{region 'Documentation'}
(*!
<summary>Check that IN is inside the inclusive StartTime..EndTime interval.</summary>
<description>

StartTime &gt; EndTime reports Error during active evaluation; equal bounds are
valid.

</description>
*)
{endregion}
FUNCTION_BLOCK AssertInTimespan_DT EXTENDS AssertionBase
VAR_INPUT
    IN : DT; //! Actual value checked or observed by this Assertion.
    StartTime : DT; //! Inclusive start of the time span; must not exceed EndTime.
    EndTime : DT; //! Inclusive end of the time span; must not precede StartTime.
END_VAR

SUPER^();

{region 'Documentation'}
(*!
<summary>Evaluate the typed temporal relation and report higher-priority errors first.</summary>
*)
{endregion}
METHOD PROTECTED Assert
VAR
    Message : STRING(GVL_Constants.MessageLength);
    StartTimeText : STRING(GVL_Constants.AssertionValueLength);
    EndTimeText : STRING(GVL_Constants.AssertionValueLength);
    ActualText : STRING(GVL_Constants.AssertionValueLength);
END_VAR
IF NOT EvaluationActive THEN
    RETURN;
END_IF;

IF Result = E_Result.Error THEN
    RETURN;
END_IF;

IF StartTime > EndTime THEN
    StartTimeText := DT_TO_STRING(StartTime);
    EndTimeText := DT_TO_STRING(EndTime);
    Message := CONCAT('Assertion error: start time exceeds end time. StartTime = ',
        StartTimeText);
    Message := CONCAT(Message, ', EndTime = ');
    Message := CONCAT(Message, EndTimeText);
    Message := CONCAT(Message, '.');
    Error(Message := Message);
    RETURN;
END_IF;

IF Result = E_Result.Failed THEN
    RETURN;
END_IF;

IF (IN < StartTime) OR (IN > EndTime) THEN
    StartTimeText := DT_TO_STRING(StartTime);
    EndTimeText := DT_TO_STRING(EndTime);
    ActualText := DT_TO_STRING(IN);
    Message := CONCAT('Assertion failed: value is outside allowed timespan. StartTime = ',
        StartTimeText);
    Message := CONCAT(Message, ', EndTime = ');
    Message := CONCAT(Message, EndTimeText);
    Message := CONCAT(Message, ', Actual = ');
    Message := CONCAT(Message, ActualText);
    Message := CONCAT(Message, '.');
    Fail(Message := Message);
    RETURN;
END_IF;

Pass();
END_METHOD

END_FUNCTION_BLOCK

(* stored: Version 1.1.0.1
   POU AssertInTimespan_DT: Id {b224fd11-3ab3-4bf6-befe-f267d3460e99}, SpecialFunc None
   Folder Internal: Id {25bc37b8-3f4e-491c-bad1-aa670c5122bc}
   Method Assert: Id {a28706ef-2fd5-4669-b958-bd1eb0803bf0} *)
